Fanuc KAREL source: KT00597.KL

PROGRAM KT00597
%NOLOCKGROUP
VAR
  R1: REAL
  R2: REAL
  OUT: STRING[80]
BEGIN
  R1 = 2.0
  R2 = 3.0
  R1 = 2.0
  R2 = 3.0
  OUT = R1 + R2
END KT00597
